(* IEC 61131-3 sources: plc-vscode/tests/st/test-ready/rusty/tests/lit/multi/pic_flags, 2 files *)

(* ---- helper.st ---- *)
FUNCTION helper : DINT
helper := 42;
END_FUNCTION

FUNCTION doubler : DINT
VAR_INPUT
    x : DINT;
END_VAR
doubler := x * 2;
END_FUNCTION

(* ---- main.st ---- *)
FUNCTION main : DINT
VAR
    result : DINT;
END_VAR
result := helper();
printf('%d$N', result);
printf('%d$N', doubler(result));
main := 0;
END_FUNCTION
